Fanuc KAREL source: KT00653.KL

PROGRAM KT00653
%NOLOCKGROUP
VAR
  P1: POSITION
  P2: POSITION
  OUT: REAL
BEGIN
  OUT = NOT P1
END KT00653
